{attribute 'linkalways'} 
{attribute 'no_explicit_call' := 'This FB is a CLASS and must be accessed using methods or properties'}
{attribute 'enable_dynamic_creation'}
FUNCTION_BLOCK _ETcVnHoughMethod EXTENDS EnumDatatypeBase
VAR
	localData : ETcVnHoughMethod;
	activeData : REFERENCE TO ETcVnHoughMethod;
	enumBaseDatatype : _DINT(localData);
END_VAR

METHOD PRIVATE AddLocalEnumeration
VAR_INPUT
	Enumeration : T_MAXSTRING;
	Value : ETcVnHoughMethod;
END_VAR
AddEnumeration(Enumeration, Value);
END_METHOD

PROPERTY PUBLIC Address : PVOID
GET
Address := ADR(activeData);
END_GET
END_PROPERTY

METHOD PUBLIC ClearReference
VAR_INPUT
END_VAR
activeData REF= localData;
SetBaseDatatypeReference();
END_METHOD

METHOD PUBLIC Clone : I_Datatype
VAR
    pClone : POINTER TO _ETcVnHoughMethod;
END_VAR
pClone := __NEW(_ETcVnHoughMethod(InitialValue := Value));
Clone := pClone^;
END_METHOD

METHOD FB_init : BOOL
VAR_INPUT
	bInitRetains : BOOL; // if TRUE, the retain variables are initialized (warm start / cold start)
	bInCopyCode : BOOL;  // if TRUE, the instance afterwards gets moved into the copy code (online change)
	InitialValue : ETcVnHoughMethod;
END_VAR
localData := InitialValue;
AddBaseDatatype(enumBaseDatatype);
ClearReference();

AddLocalEnumeration('TCVN_HM_STANDARD', ETcVnHoughMethod.TCVN_HM_STANDARD);
AddLocalEnumeration('TCVN_HM_PROBABILISTIC', ETcVnHoughMethod.TCVN_HM_PROBABILISTIC);
AddLocalEnumeration('TCVN_HM_MULTI_SCALE', ETcVnHoughMethod.TCVN_HM_MULTI_SCALE);
AddLocalEnumeration('TCVN_HM_GRADIENT', ETcVnHoughMethod.TCVN_HM_GRADIENT);
AddLocalEnumeration('TCVN_HM_GRADIENT_ALT', ETcVnHoughMethod.TCVN_HM_GRADIENT_ALT);
END_METHOD

PROPERTY PUBLIC Identifier : T_MAXSTRING
GET
Identifier := 'ETcVnHoughMethod';
END_GET
END_PROPERTY

METHOD IsEnumeratorValueEqual : BOOL
VAR_INPUT
	Enumerator : I_KeyValueForwardEnumerator;
END_VAR
VAR
	storedValue : ETcVnHoughMethod;
END_VAR
IF NOT Enumerator.TryGet(storedValue) THEN
	RETURN;
END_IF

IsEnumeratorValueEqual := storedValue = activeData;
END_METHOD

METHOD PUBLIC MakeReferenceTo
VAR_INPUT
	ReferenceTarget : REFERENCE TO ETcVnHoughMethod;
END_VAR
activeData REF= ReferenceTarget;
SetBaseDatatypeReference();
END_METHOD

METHOD PROTECTED SetBaseDatatypeReference
VAR_INPUT
END_VAR
enumBaseDatatype.MakeReferenceTo(activeData);
END_METHOD

PROPERTY PUBLIC Size : UDINT
GET
Size := SIZEOF(activeData);
END_GET
END_PROPERTY

METHOD TryMakeReferenceTo : BOOL
VAR_INPUT
	Target : I_Datatype;
END_VAR
VAR
	pTargetData : POINTER TO ETcVnHoughMethod;
END_VAR
IF NOT IsEquivalentTo(Target) THEN
	RETURN;
END_IF

pTargetData := Target.Address;
activeData REF= pTargetData^;
SetBaseDatatypeReference();
TryMakeReferenceTo := TRUE;
END_METHOD

PROPERTY PUBLIC Value : ETcVnHoughMethod
GET
Value := activeData;
END_GET
SET
activeData := Value;
END_SET
END_PROPERTY

END_FUNCTION_BLOCK

(* stored: Version 1.1.0.1, ProductVersion 3.1.4024.13
   POU _ETcVnHoughMethod: Id {8e8e81ba-7bc2-0eb0-0aa6-b932849bfacf}, SpecialFunc None
   Folder Core: Id {ed0f5fa3-4a79-0ae9-166d-a8cebb75ec22}
   Folder Protected: Id {2e28e7a6-7637-0b2c-08f6-2e6eaca4ac2a}
   Folder Customize: Id {7735d64d-94a8-004e-1a7b-20f832eeb266}
   Folder Constructor: Id {825a3143-73ff-0ac0-1490-f66c3f30edf0}
   Folder Private: Id {2d7bfa7f-af78-0d27-2806-91775ddc4d78}
   Folder Protected: Id {9b798fd3-90ae-05b0-365e-a1b98ad5af53}
   Method AddLocalEnumeration: Id {d594f1db-523a-018c-35d2-fa9c98b06a13}
   Property Address: Id {a1877ceb-7d5d-0ef4-2634-b2e2c982a19e}
   Get Get: Id {70bcfd3d-ab00-0d7f-2c3e-f15614b8a556}
   Method ClearReference: Id {04d0bfa2-e550-0d69-301f-b05614911280}
   Method Clone: Id {99b9c5a2-4592-00ba-38be-70f77148bf5b}
   Method FB_init: Id {85b8c148-50be-0f3c-04f1-9ec00b42c47f}
   Property Identifier: Id {ef6a9525-e29a-0146-3570-b249750796a0}
   Get Get: Id {4995b785-da1d-0562-2a96-340aa0c394cf}
   Method IsEnumeratorValueEqual: Id {0ff8d33d-0455-07cd-2d8b-48bbe6103a14}
   Method MakeReferenceTo: Id {61e4f5fd-7d7a-0ac8-0856-88fe62fb6b54}
   Method SetBaseDatatypeReference: Id {0c86be6f-2a98-0f48-0ee5-1ef46e2aad24}
   Property Size: Id {65a0766a-f46c-05ae-2727-54f829180e31}
   Get Get: Id {28564351-b385-0770-1e21-ca24357cb67d}
   Method TryMakeReferenceTo: Id {08816ede-525c-04d5-01e3-a256f8c9ca83}
   Property Value: Id {4d0326cc-7d48-044c-2c2a-505c12523b9f}
   Get Get: Id {376be4ff-3d15-09b4-3279-0d0e093ce550}
   Set Set: Id {f0803f8a-a67e-0d4c-0817-2ced4c3c41d7} *)
